(* IEC 61131-3 sources: ZPLC/packages/zplc-ide/projects/kitchen_sink/src, 10 files *)

(* ---- bits_scaling.st ---- *)
(*
 * Kitchen Sink 6/10 - bitwise, logic, conversion, scaling and system functions
 *
 * SPDX-License-Identifier: MIT
 *)

PROGRAM KsBitsScaling
VAR
    StartButton     : BOOL := FALSE;
    StopButton      : BOOL := FALSE;
    SensorInput     : REAL := 50.0;
    TempBool        : BOOL;
    TempInt         : INT := 0;
    TempReal        : REAL := 0.0;
    Normalized      : REAL := 0.0;
    Scaled          : REAL := 0.0;
    SysUptime       : DINT := 0;
    SysCycleTime    : DINT := 0;
END_VAR

(* ============================================================================
 * SECTION 11: Bitwise Functions
 * ============================================================================ *)

TempInt := SHL(1, 4);       (* 1 << 4 = 16 *)
TempInt := SHR(256, 4);     (* 256 >> 4 = 16 *)
TempInt := ROL(1, 31);      (* Rotate left *)
TempInt := ROR(1, 1);       (* Rotate right *)

(* ============================================================================
 * SECTION 12: Logic Functions
 * ============================================================================ *)

TempBool := NAND(StartButton, StopButton);
TempBool := NOR(StartButton, StopButton);

(* ============================================================================
 * SECTION 13: Type Conversion Functions
 * ============================================================================ *)

TempReal := INT_TO_REAL(TempInt);
TempInt := REAL_TO_INT(TempReal);
TempInt := BOOL_TO_INT(StartButton);
TempBool := INT_TO_BOOL(TempInt);

(* ============================================================================
 * SECTION 14: Scaling Functions
 * ============================================================================ *)

Normalized := NORM_X(0.0, SensorInput, 100.0);
Scaled := SCALE_X(0.0, Normalized, 4095.0);

(* ============================================================================
 * SECTION 15: System Functions
 * ============================================================================ *)

SysUptime := UPTIME();
SysCycleTime := CYCLE_TIME();
WATCHDOG_RESET();

END_PROGRAM

(* ---- buffers.st ---- *)
(*
 * Kitchen Sink 4/10 - system buffer blocks
 *
 * Blocks: FIFO, LIFO (64 and 56 bytes with the default SIZE of 8). As in the
 * original fixture they are declared, which allocates them, but never called.
 *
 * SPDX-License-Identifier: MIT
 *)

PROGRAM KsBuffers
VAR
    FifoBuffer      : FIFO;
    LifoBuffer      : LIFO;
END_VAR

END_PROGRAM

(* ---- math.st ---- *)
(*
 * Kitchen Sink 5/10 - selection, math, trigonometry and logarithm functions
 *
 * SPDX-License-Identifier: MIT
 *)

PROGRAM KsMath
VAR
    SensorInput     : REAL := 50.0;
    SelectFlag      : BOOL := FALSE;
    TempInt         : INT := 0;
    TempReal        : REAL := 0.0;
    Angle           : REAL := 0.785398; (* PI/4 = 45 degrees *)
END_VAR

(* ============================================================================
 * SECTION 7: Selection Functions
 * ============================================================================ *)

TempReal := MAX(SensorInput, 25.0);
TempReal := MIN(TempReal, 75.0);
TempReal := LIMIT(0.0, SensorInput, 100.0);
TempReal := SEL(SelectFlag, 0.0, SensorInput);
TempInt := MUX(1, 10, 20, 30);

(* ============================================================================
 * SECTION 8: Math Functions
 * ============================================================================ *)

TempReal := ABS(-42.5);
TempInt := ABS(-100);
TempReal := NEG(SensorInput);
TempInt := 17 MOD 5;        (* MOD is an infix operator in IEC 61131-3 *)
TempReal := SQRT(144.0);
TempReal := EXPT(2.0, 8.0);
TempReal := TRUNC(3.7);
TempReal := ROUND(3.5);

(* ============================================================================
 * SECTION 9: Trigonometry Functions
 * ============================================================================ *)

TempReal := SIN(Angle);
TempReal := COS(Angle);
TempReal := TAN(Angle);
TempReal := ASIN(0.5);
TempReal := ACOS(0.5);
TempReal := ATAN(1.0);
TempReal := ATAN2(1.0, 1.0);

(* ============================================================================
 * SECTION 10: Logarithmic Functions
 * ============================================================================ *)

TempReal := LN(2.718281828);
TempReal := LOG(100.0);
TempReal := EXP(1.0);

END_PROGRAM

(* ---- pid.st ---- *)
(*
 * Kitchen Sink 3/10 - PID controller
 *
 * Block: PID_Compact (48 bytes of instance data, so it gets a program of its
 * own), plus LIMIT on its output.
 *
 * SPDX-License-Identifier: MIT
 *)

PROGRAM KsPid
VAR
    SensorInput     : REAL := 50.0;
    AnalogOutput    : REAL := 0.0;
    TempReal        : REAL := 0.0;
    PidController   : PID_Compact;
END_VAR

(* PID_Compact - PID Controller *)
(* KI is KP / TI and KD is KP * TD in the units of the block; DT is the sample time in seconds *)
PidController(
    SP := 50.0,
    PV := SensorInput,
    KP := 1.0,
    KI := 1.0,
    KD := 0.1,
    DT := 0.01,
    OUT_MIN := 0.0,
    OUT_MAX := 100.0
);

TempReal := LIMIT(0.0, PidController.OUT, 100.0);
AnalogOutput := LIMIT(0.0, PidController.OUT, 100.0);

END_PROGRAM

(* ---- process_control.st ---- *)
(*
 * Kitchen Sink 2/10 - process control blocks
 *
 * Blocks: HYSTERESIS, DEADBAND, LAG_FILTER, RAMP_REAL, INTEGRAL, DERIVATIVE
 * (PID_Compact has its own program, pid.st: it alone takes 48 bytes.)
 *
 * SPDX-License-Identifier: MIT
 *)

PROGRAM KsProcess
VAR
    (* ===== Inputs ===== *)
    SensorInput     : REAL := 50.0;
    StopButton      : BOOL := FALSE;

    (* ===== Outputs ===== *)
    MotorPermit     : BOOL := FALSE;

    (* ===== Process Control FBs ===== *)
    HystCtrl        : HYSTERESIS;
    DeadCtrl        : DEADBAND;
    LagFilt         : LAG_FILTER;
    RampCtrl        : RAMP_REAL;
    Integrator      : INTEGRAL;
    Differentiator  : DERIVATIVE;
END_VAR

(* HYSTERESIS - On/Off control with deadband *)
HystCtrl(IN := SensorInput, HIGH := 60.0, LOW := 40.0);

(* DEADBAND - Filter small changes *)
DeadCtrl(IN := SensorInput, WIDTH := 2.0);

(* LAG_FILTER - First-order lag filter *)
(* GAIN is the share of the difference taken each scan: 10 ms / (100 ms + 10 ms) *)
LagFilt(IN := SensorInput, GAIN := 0.09);

(* RAMP_REAL - Rate limiter *)
RampCtrl(IN := SensorInput, RATE := 10.0);

(* INTEGRAL - Integration *)
(* DT is the sample time in seconds *)
Integrator(IN := 1.0, DT := 0.01, RESET := StopButton);

(* DERIVATIVE - Differentiation *)
Differentiator(IN := SensorInput, DT := 0.01);

(* Final output: the motor is allowed only while the sensor is not above HIGH *)
MotorPermit := NOT HystCtrl.Q;

END_PROGRAM

(* ---- sequencing.st ---- *)
(*
 * Kitchen Sink 1/10 - timers, edges, bistables, counters, generators
 *
 * Part of the standard-library conformance fixture. The original single
 * program needed about 770 bytes of WORK memory, but every PROGRAM owns a
 * 256-byte region (WORK_MEMORY_REGION_SIZE, init flag included), so the
 * fixture is split into ten small programs, one per task. Each program
 * keeps the blocks that feed each other together.
 *
 * Blocks: TON, TOF, TP, R_TRIG, F_TRIG, RS, SR, CTU, CTD, CTUD, BLINK, PWM, PULSE
 *
 * SPDX-License-Identifier: MIT
 *)

PROGRAM KsSequencing
VAR
    (* ===== Inputs ===== *)
    StartButton     : BOOL := FALSE;
    StopButton      : BOOL := FALSE;
    CounterPulse    : BOOL := FALSE;

    (* ===== Outputs ===== *)
    MotorOutput     : BOOL := FALSE;
    AlarmOutput     : BOOL := FALSE;

    (* ===== Timer FBs ===== *)
    TimerOn         : TON;
    TimerOff        : TOF;
    TimerPulse      : TP;

    (* ===== Edge Detection FBs ===== *)
    RisingEdge      : R_TRIG;
    FallingEdge     : F_TRIG;

    (* ===== Bistable FBs ===== *)
    Latch_RS        : RS;
    Latch_SR        : SR;

    (* ===== Counter FBs ===== *)
    CountUp         : CTU;
    CountDown       : CTD;
    CountUpDown     : CTUD;

    (* ===== Generator FBs ===== *)
    Blinker         : BLINK;
    PwmGen          : PWM;
    PulseGen        : PULSE;
END_VAR

(* ============================================================================
 * SECTION 1: Timer Function Blocks
 * ============================================================================ *)

(* TON - On-delay timer *)
TimerOn(IN := StartButton, PT := T#1000ms);

(* TOF - Off-delay timer *)
TimerOff(IN := TimerOn.Q, PT := T#500ms);

(* TP - Pulse timer *)
TimerPulse(IN := StopButton, PT := T#200ms);

(* ============================================================================
 * SECTION 2: Edge Detection
 * ============================================================================ *)

(* R_TRIG - Rising edge detection *)
RisingEdge(CLK := StartButton);

(* F_TRIG - Falling edge detection *)
FallingEdge(CLK := StopButton);

(* ============================================================================
 * SECTION 3: Bistable Latches
 * ============================================================================ *)

(* RS - Reset-dominant latch *)
Latch_RS(S := RisingEdge.Q, R1 := FallingEdge.Q);

(* SR - Set-dominant latch *)
Latch_SR(S1 := RisingEdge.Q, R := FallingEdge.Q);

(* ============================================================================
 * SECTION 4: Counters
 * ============================================================================ *)

(* CTU - Count Up *)
CountUp(CU := CounterPulse, R := StopButton, PV := 100);

(* CTD - Count Down *)
CountDown(CD := CounterPulse, LD := StartButton, PV := 50);

(* CTUD - Count Up/Down *)
CountUpDown(CU := RisingEdge.Q, CD := FallingEdge.Q, R := StopButton, LD := FALSE, PV := 200);

(* ============================================================================
 * SECTION 5: Generators
 * ============================================================================ *)

(* BLINK - Oscillator *)
Blinker(ENABLE := Latch_RS.Q1, T_ON := T#500ms, T_OFF := T#500ms);

(* PWM - Pulse Width Modulation *)
PwmGen(ENABLE := TRUE, PERIOD := T#1000ms, DUTY := 75);

(* PULSE - Single pulse generator *)
PulseGen(TRIG := RisingEdge.Q, PT := T#100ms);

(* ============================================================================
 * SECTION 6: Outputs
 * ============================================================================ *)

MotorOutput := Latch_RS.Q1 AND TimerOff.Q;
AlarmOutput := CountUp.Q OR Blinker.Q;

END_PROGRAM

(* ---- strings_build.st ---- *)
(*
 * Kitchen Sink 8/10 - string functions, part 2 (join and cut)
 *
 * Functions: CONCAT, LEFT, RIGHT, MID
 *
 * SPDX-License-Identifier: MIT
 *)

PROGRAM KsStringsBuild
VAR
    Str1            : STRING := 'Hello';
    StrResult       : STRING;
END_VAR

StrResult := CONCAT(Str1, ' ');
StrResult := CONCAT(StrResult, 'World');
StrResult := LEFT(Str1, 3);
StrResult := RIGHT(StrResult, 3);
StrResult := MID(Str1, 2, 3);

END_PROGRAM

(* ---- strings_compare.st ---- *)
(*
 * Kitchen Sink 10/10 - string functions, part 4 (copy and compare)
 *
 * Functions: COPY, STRCMP, EQ_STRING, NE_STRING
 *
 * SPDX-License-Identifier: MIT
 *)

PROGRAM KsStringsCompare
VAR
    Str1            : STRING := 'Hello';
    Str2            : STRING := 'World';
    TempInt         : INT := 0;
    TempBool        : BOOL;
END_VAR

Str2 := COPY(Str1, Str2);        (* COPY(src, dst) returns dst *)
TempInt := STRCMP(Str1, Str2);
TempBool := EQ_STRING(Str1, 'Hello');
TempBool := NE_STRING(Str1, Str2);

END_PROGRAM

(* ---- strings_edit.st ---- *)
(*
 * Kitchen Sink 9/10 - string functions, part 3 (edit)
 *
 * Functions: INSERT, DELETE, REPLACE, CLEAR
 *
 * SPDX-License-Identifier: MIT
 *)

PROGRAM KsStringsEdit
VAR
    Str1            : STRING := 'Hello';
    StrResult       : STRING;
END_VAR

StrResult := INSERT(Str1, '!!!', 5);
StrResult := DELETE(StrResult, 3, 5);
StrResult := REPLACE(Str1, 'Hi', 1, 2);
StrResult := CLEAR(StrResult);   (* CLEAR returns the cleared string *)

END_PROGRAM

(* ---- strings_measure.st ---- *)
(*
 * Kitchen Sink 7/10 - string functions, part 1 (measure)
 *
 * A STRING takes 85 bytes of the program's 256-byte WORK region and string
 * literals live there too, so the string functions are spread over four
 * programs with at most two STRING variables each.
 *
 * Functions: LEN, FIND
 *
 * SPDX-License-Identifier: MIT
 *)

PROGRAM KsStringsMeasure
VAR
    Str1            : STRING := 'Hello';
    StrLen          : INT := 0;
    StrPos          : INT := 0;
END_VAR

StrLen := LEN(Str1);
StrPos := FIND(Str1, 'ell');

END_PROGRAM
